Fanuc KAREL source: ko00047.KL

-- PROVISIONAL review KL for V1013-1; original PC SHA256 787a58ee353c187ae8a732533e80a9b2367c86a36025f4fdf3095b46f86abcf6
-- Incomplete behavior may be omitted. Consult companion uncertainty JSON. Do not deploy.
PROGRAM KO00047
%NOLOCKGROUP
BEGIN
  -- UNRESOLVED_PC offsets 5-12; opcodes 9D,23
  -- UNRESOLVED_PC offsets 17-69; opcodes 27,27,49,7E,AD,27,49,7E,AD,22,31,7E,4A
  -- UNRESOLVED_PC offsets 74-78; opcodes 7F
END KO00047
